(* IEC 61131-3 sources: Test-Git_ESME26/TestProgettoESME_26.fbsproj/PacDriveLib Migration/Motion/Homing (part 2) *)

(* ---- PDL_FB_HomeSetPos.fb.st ---- *)
FUNCTION_BLOCK PDL_FB_HomeSetPos
VAR_INPUT
	i_xEnable             : BOOL;
	i_ifDrive             : MOIN.IF_Axis;
	i_etMode              : PDL_ET_HomeSetPosMode;
	i_lrHomePosition      : LREAL;
	i_lrEncoderPosition   : LREAL;
	i_lrAbsEncOffset      : LREAL;
	i_lrUserPeriod        : LREAL;
	i_lrRestoreWindow     : LREAL;
	i_pstRestorePosRetain : POINTER TO PDL_ST_AxisRestorePosition;
	i_xExecute            : BOOL;
	iq_lencEncoder        : MOIN.IF_LogicalEncoder;
END_VAR
VAR_OUTPUT
	q_xActive           : BOOL;
	q_xReady            : BOOL;
	q_xBusy             : BOOL;
	q_xDone             : BOOL;
	q_etDiag            : GD.ET_Diag     := GD.ET_Diag.Ok;
	q_etDiagExt         : PDL_ET_DiagExt := PDL_ET_DiagExt.Disabled;
	q_sMsg              : STRING[80];
	q_lrPosition        : LREAL;
	q_lrEncoderPosition : LREAL;
	q_xHomeOk           : BOOL;
END_VAR
VAR
	xEnableFlag                                : BOOL;
	diState                                    : DINT;
	lrEncoderPeriode                           : LREAL;
	lrTurns                                    : LREAL;
	lrModuloPosition                           : LREAL;
	lrEncPosition                              : LREAL;
	xInterfacesInitialized                     : BOOL;
	xSuccess                                   : BOOL;
	etDiagTemp                                 : GD.ET_Diag := GD.ET_Diag.Ok;
	etDiagExtTemp                              : PDL_ET_DiagExt := PDL_ET_DiagExt.Ok;
	sDummyString                               : STRING[80];
	fbLoggerPoint                              : APL.FB_LoggerPoint;
	fbSetPosAxis                               : PLCO.MC_SetPosition;
	fbSetPosLenc                               : PLCO.MC_SetPosition;
	ifScalingAccess                            : DMFI.IF_ScalingAccess;
	ifScaling                                  : DMFI.IF_Scaling;
	ifGetParentDevice                          : DTSI.IF_GetParentDevice;
	ifDeviceAccess                             : DTSI.IF_DeviceAccess;
	ifEncoderAccess                            : DDI.IF_EncoderAccess;
	ifEncoder                                  : DDI.IF_Encoder;
	etModeOld                                  : PDL_ET_HomeSetPosMode;
	lrQuotientEncPeriodToUserPeriod            : LREAL;
	diTruncFromQuotient                        : DINT;
	lrAbsDifferenceQuotientToTruncFromQuotient : LREAL;
	xUserPeriodFitsIntoEncoderPeriod           : BOOL;
END_VAR

IF i_xEnable AND NOT xEnableFlag THEN (* Input action by rising edge of enable *)
	xEnableFlag := TRUE;
	THIS^.fbLoggerPoint.AddLogEntry(
		i_etLogLevel := APL.ET_LogLevel.UserAction, i_etDiag := q_etDiag, i_udiDiagExt := q_etDiagExt, i_sMessage := 'enable function block',
	);
	q_xActive              := TRUE;
	q_xReady               := FALSE;
	q_xBusy                := FALSE;
	q_xDone                := FALSE;
	q_xHomeOk              := FALSE;
	xInterfacesInitialized := Init_Interfaces();
	IF xInterfacesInitialized THEN
		etModeOld := i_etMode;
		q_xReady  := TRUE;
		SetDiagOutput(i_etDiag := GD.ET_Diag.OK, i_etDiagExt := PDL_ET_DiagExt.WaitForExecute, i_sMsg := '');
		diState := 10;
	END_IF
	i_ifDrive.xIsHomed := FALSE;

ELSIF NOT i_xEnable AND xEnableFlag THEN (* Output action by falling edge of enable *)
	xEnableFlag := FALSE;
	THIS^.fbLoggerPoint.AddLogEntry(
		i_etLogLevel := APL.ET_LogLevel.UserAction, i_etDiag := q_etDiag, i_udiDiagExt := q_etDiagExt, i_sMessage := 'disable function block',
	);
	xInterfacesInitialized := FALSE;
	q_xActive              := FALSE;
	q_xReady               := FALSE;
	q_xBusy                := FALSE;
	q_xDone                := FALSE;
	q_lrPosition           := 0.0;
	q_lrEncoderPosition    := 0.0;
	q_xHomeOk              := FALSE;
	SetDiagOutput(i_etDiag := GD.ET_Diag.Ok, i_etDiagExt := PDL_ET_DiagExt.Disabled, i_sMsg := '');
	diState := 0;
ELSIF NOT q_xActive THEN
	RETURN;
END_IF

IF xInterfacesInitialized THEN
	q_lrPosition        := i_ifDrive.RefPosition;
	IF iq_lencEncoder <> 0 THEN
		q_lrEncoderPosition := iq_lencEncoder.RefPosition;
	ELSE
		q_lrEncoderPosition := 0;
	END_IF
	q_xBusy             := q_etDiag = GD.ET_Diag.Ok AND NOT q_xDone AND diState > 10;
ELSE
	diState  := 0;
	q_xReady := FALSE;
	RETURN;
END_IF

CASE diState OF
	0: (* Idle *)
		;
	10: (* wait for xExecute *)
		IF i_xExecute THEN
			IF etModeOld <> i_etMode THEN
				etModeOld              := i_etMode;
				xInterfacesInitialized := Init_Interfaces();
			END_IF
			lrEncoderPeriode := 0;

			THIS^.fbLoggerPoint.AddLogEntry(
				i_etLogLevel := APL.ET_LogLevel.UserAction,
				i_etDiag     := q_etDiag,
				i_udiDiagExt := q_etDiagExt,
				i_sMessage   := 'start homing',
				q_etDiag     =>,
				q_etDiagExt  =>
			);

			lrEncoderPeriode 			:= ifEncoder.Revolutions
											* ifScaling.PositionResolution
											* TO_LREAL(ifScaling.GearIn) / TO_LREAL(ifScaling.GearOut)
											* TO_LREAL( ifEncoder.GearOut) / TO_LREAL(ifEncoder.GearIn);

						// Calculation if UserPeriod fits into EncoderPeriod
			IF (i_lrUserPeriod > CMT.Gc_lrZeroTolerance) AND (lrEncoderPeriode > CMT.Gc_lrZeroTolerance) THEN

				lrQuotientEncPeriodToUserPeriod					:= lrEncoderPeriode/i_lrUserPeriod;
				diTruncFromQuotient 							:= TRUNC(lrQuotientEncPeriodToUserPeriod);
				lrAbsDifferenceQuotientToTruncFromQuotient		:= ABS (lrQuotientEncPeriodToUserPeriod - TO_LREAL(diTruncFromQuotient));

				IF (lrAbsDifferenceQuotientToTruncFromQuotient < CMT.Gc_lrZeroTolerance)
				OR ((1 - lrAbsDifferenceQuotientToTruncFromQuotient < CMT.Gc_lrZeroTolerance) AND (lrAbsDifferenceQuotientToTruncFromQuotient <= 1)) THEN
					xUserPeriodFitsIntoEncoderPeriod	:= TRUE;
				ELSE
					xUserPeriodFitsIntoEncoderPeriod	:= FALSE;
				END_IF

			END_IF

			CASE i_etMode OF
				//---------------------------------------
				PDL_ET_HomeSetPosMode.RestorePosFromRetain,
				PDL_ET_HomeSetPosMode.SetPosAxisPosition,
				PDL_ET_HomeSetPosMode.SetPosLogEncoderPosition,
				PDL_ET_HomeSetPosMode.SetPosAxisAndLogEncoderPosition,
				PDL_ET_HomeSetPosMode.RestorePosFromAxisencoder:
					//---------------------------------------

					//Input-Parameter-Checks
					IF i_etMode = PDL_ET_HomeSetPosMode.RestorePosFromAxisEncoder OR i_etMode = PDL_ET_HomeSetPosMode.RestorePosFromRetain THEN
						IF (ABS(ifEncoder.Revolutions) < 1.0E-3) THEN
							SetDiagOutput(	i_etDiag := GD.ET_Diag.DriveConditionInvalid,
											i_etDiagExt := PDL_ET_DiagExt.DriveEncoderInvalid,
											i_sMsg := ''
							);
							diState := 0;
							RETURN;
						END_IF

						IF (i_lrUserPeriod < 0.0) THEN
							SetDiagOutput(
								i_etDiag    := GD.ET_Diag.InputParameterInvalid,
								i_etDiagExt := PDL_ET_DiagExt.UserPeriodRange,
								i_sMsg      := '0.0 <= i_lrUserPeriod'
							);
							diState := 0;
							RETURN;
							// if UserPeriod = 0: Check if AbsEncOffset > 0
						ELSIF
							i_etMode = PDL_ET_HomeSetPosMode.RestorePosFromAxisencoder AND
							(i_lrUserPeriod = 0.0) AND
							((i_lrAbsEncOffset < 0) OR (i_lrAbsEncOffset > lrEncoderPeriode))
						THEN
							SetDiagOutput(
								i_etDiag    := GD.ET_Diag.InputParameterInvalid,
								i_etDiagExt := PDL_ET_DiagExt.AbsEncOffsetRange,
								i_sMsg      := STANDARD.CONCAT('0.0 < i_lrAbsEncOffset <= ', SE_CTBX.FC_LrealToString(i_sFormat := '#0.00', i_lrInput := lrEncoderPeriode))
							);
							diState := 0;
							RETURN;
							// Check if UserPeriode fits into EncoderPeriode
						ELSIF i_etMode = PDL_ET_HomeSetPosMode.RestorePosFromAxisencoder AND (i_lrUserPeriod > 0.0) AND NOT xUserPeriodFitsIntoEncoderPeriod
						THEN
							SetDiagOutput(
								i_etDiag    := GD.ET_Diag.InputParameterInvalid,
								i_etDiagExt := PDL_ET_DiagExt.UserPeriodRange,
								i_sMsg      := STANDARD.CONCAT('i_lrUserPeriod has to be a divsior of ',SE_CTBX.FC_LrealToString(i_sFormat := '#0.00', i_lrInput := lrEncoderPeriode))
							);
							diState := 0;
							RETURN;
						END_IF
					END_IF

					q_xHomeOk := FALSE;
					q_xBusy   := TRUE;
					q_xDone   := FALSE;
					SetDiagOutput(i_etDiag := GD.ET_Diag.Ok, i_etDiagExt := PDL_ET_DiagExt.WaitUntilHomingDone, i_sMsg := '');
					diState := 20;
				ELSE
					SetDiagOutput(i_etDiag := GD.ET_Diag.InputParameterInvalid, i_etDiagExt := PDL_ET_DiagExt.UnknownMode, i_sMsg := '');
					diState := 0;
			END_CASE
		END_IF
	20:
		CASE i_etMode OF
			//---------------------------------------
			PDL_ET_HomeSetPosMode.RestorePosFromRetain: (* Restore axis position from stored and actual Values of position and encoder position *)
				//---------------------------------------
				IF i_pstRestorePosRetain > 0 THEN
					PDL_FC_RestoreAxisPosition(
						i_ifDrive           := i_ifDrive,
						i_lrUserPeriod      := i_lrUserPeriod,
						i_lrRestoreWindow   := i_lrRestoreWindow,
						i_stRestorePosition := i_pstRestorePosRetain^,
						q_etDiag            => etDiagTemp,
						q_etDiagExt         => etDiagExtTemp,
						q_sMsg              => sDummyString
					);
					IF etDiagTemp = GD.ET_Diag.Ok THEN
						diState := 30;
					ELSE
						CASE etDiagExtTemp OF
							PDL_ET_DiagExt.CheckSumInvalid:
								SetDiagOutput(
									i_etDiag    := GD.ET_Diag.InputParameterInvalid,
									i_etDiagExt := PDL_ET_DiagExt.CheckSumInvalid,
									i_sMsg      := 'FB_HomeSetPos: FC_RestoreAxisPosition'
								);
							PDL_ET_DiagExt.DataNVRamInvalid:
								SetDiagOutput(
									i_etDiag    := GD.ET_Diag.InputParameterInvalid,
									i_etDiagExt := PDL_ET_DiagExt.DataNVRamInvalid,
									i_sMsg      := 'FB_HomeSetPos: FC_RestoreAxisPosition'
								);
							PDL_ET_DiagExt.SercosNotInPhaseFour:
								SetDiagOutput(
									i_etDiag    := GD.ET_Diag.DriveConditionInvalid,
									i_etDiagExt := PDL_ET_DiagExt.SercosNotInPhaseFour,
									i_sMsg      := 'FB_HomeSetPos: FC_RestoreAxisPosition'
								);
							PDL_ET_DiagExt.DriveEncoderInvalid:
								SetDiagOutput(
									i_etDiag    := GD.ET_Diag.DriveConditionInvalid,
									i_etDiagExt := PDL_ET_DiagExt.DriveEncoderInvalid,
									i_sMsg      := 'FB_HomeSetPos: FC_RestoreAxisPosition'
								);
							PDL_ET_DiagExt.OutOfRestoreWindow:
								SetDiagOutput(
									i_etDiag    := GD.ET_Diag.LimitReached,
									i_etDiagExt := PDL_ET_DiagExt.OutOfRestoreWindow,
									i_sMsg      := 'FB_HomeSetPos: FC_RestoreAxisPosition'
								);
							PDL_ET_DiagExt.UnexpectedFeedback:
								SetDiagOutput(
									i_etDiag    := GD.ET_Diag.UnexpectedProgramBehavior,
									i_etDiagExt := PDL_ET_DiagExt.UnexpectedFeedback,
									i_sMsg      := Standard.CONCAT('FB_HomeSetPos: FC_RestoreAxisPosition: ', sDummyString)
								);
							PDL_ET_DiagExt.RestoreInterrupted:
								SetDiagOutput(
									i_etDiag    := GD.ET_Diag.DriveConditionInvalid,
									i_etDiagExt := PDL_ET_DiagExt.RestoreInterrupted,
									i_sMsg      := 'FB_HomeSetPos: FC_RestoreAxisPosition'
								);
						END_CASE
						diState := 0;
					END_IF
				ELSE
					SetDiagOutput(
						i_etDiag := GD.ET_Diag.InputParameterInvalid, i_etDiagExt := PDL_ET_DiagExt.PointerRestorePosRetainInvalid, i_sMsg := ''
					);
					diState := 0;
				END_IF
				//-------------------------------------
			PDL_ET_HomeSetPosMode.SetPosAxisPosition:
				//-------------------------------------

				THIS^.fbSetPosAxis(Axis := i_ifDrive, Execute := TRUE, Position := i_lrHomePosition, Relative := FALSE);

				IF THIS^.fbSetPosAxis.Done THEN
					diState := 30;
				ELSIF THIS^.fbSetPosAxis.Error THEN
					SetDiagOutput(
						i_etDiag    := GD.ET_Diag.UnexpectedProgramBehavior,
						i_etDiagExt := PDL_ET_DiagExt.UnexpectedFeedback,
						i_sMsg      := CONCAT('MC_Setposition.ErrorID: ', PLCO.FC_EtResultToString(THIS^.fbSetPosAxis.ErrorId))
					);
					THIS^.fbSetPosAxis(Execute := FALSE);
					diState := 0;
				END_IF

				//-------------------------------------------
			PDL_ET_HomeSetPosMode.SetPosLogEncoderPosition:
				//-------------------------------------------
				THIS^.fbSetPosLenc(Axis := iq_lencEncoder, Execute := TRUE, Position := i_lrEncoderPosition, Relative := FALSE);

				IF THIS^.fbSetPosLenc.Done THEN
					diState := 30;
				ELSIF THIS^.fbSetPosLenc.Error THEN
					SetDiagOutput(
						i_etDiag    := GD.ET_Diag.UnexpectedProgramBehavior,
						i_etDiagExt := PDL_ET_DiagExt.UnexpectedFeedback,
						i_sMsg      := CONCAT('MC_Setposition.ErrorID: ', PLCO.FC_EtResultToString(THIS^.fbSetPosLenc.ErrorId))
					);
					THIS^.fbSetPosLenc(Execute := FALSE);
					diState := 0;
				END_IF

				//--------------------------------------------------
			PDL_ET_HomeSetPosMode.SetPosAxisAndLogEncoderPosition:
				//--------------------------------------------------
				THIS^.fbSetPosLenc(Axis := iq_lencEncoder, Execute := TRUE, Position := i_lrEncoderPosition, Relative := FALSE);

				THIS^.fbSetPosAxis(Axis := i_ifDrive, Execute := TRUE, Position := i_lrHomePosition, Relative := FALSE);

				IF THIS^.fbSetPosAxis.Done AND THIS^.fbSetPosLenc.Done THEN
					diState := 30;
				ELSIF THIS^.fbSetPosAxis.Error THEN
					SetDiagOutput(
						i_etDiag    := GD.ET_Diag.UnexpectedProgramBehavior,
						i_etDiagExt := PDL_ET_DiagExt.UnexpectedFeedback,
						i_sMsg      := CONCAT('MC_Setposition.ErrorID: ', PLCO.FC_EtResultToString(THIS^.fbSetPosAxis.ErrorId))
					);
					THIS^.fbSetPosAxis(Execute := FALSE);
					THIS^.fbSetPosLenc(Execute := FALSE);
					diState := 0;

				ELSIF THIS^.fbSetPosLenc.Error THEN
					SetDiagOutput(
						i_etDiag    := GD.ET_Diag.UnexpectedProgramBehavior,
						i_etDiagExt := PDL_ET_DiagExt.UnexpectedFeedback,
						i_sMsg      := CONCAT('MC_Setposition.ErrorID: ', PLCO.FC_EtResultToString(THIS^.fbSetPosLenc.ErrorId))
					);
					THIS^.fbSetPosLenc(Execute := FALSE);
					THIS^.fbSetPosAxis(Execute := FALSE);
					diState := 0;
				END_IF

				//--------------------------------------------
			PDL_ET_HomeSetPosMode.RestorePosFromAxisencoder: (* Gebertyp feststellen und GeberPeriode berechnen *)
				//--------------------------------------------
				lrTurns          := ifEncoder.Revolutions;
				IF NOT ifScaling.InvertDirection THEN (* motor direction right *)
					lrEncPosition := ifEncoder.Position;
				ELSE
					lrEncPosition := lrEncoderPeriode - ifEncoder.Position;
				END_IF
				(* In a round axis, position is always within the user period, AbsEncOffset is not allowed *)
				IF i_lrUserPeriod > 0.0 THEN
					lrModuloPosition := lrEncPosition - TRUNC_INT(lrEncPosition / i_lrUserPeriod) * i_lrUserPeriod;
					THIS^.fbSetPosAxis(Axis := i_ifDrive, Execute := TRUE, Position := lrModuloPosition, Relative := FALSE);
				ELSE
					(* Absolute axis *)
					(*---------------*)
					(* The range of the encoder period is between 0 and encoder period *)
					(* In absolute systems it makes sense to have an Offset to have neg. positions *)
					(* Of course, the Offset reduces the upper limit of the max. travel *)

					(* without AbsEncOffset *)
					(* 		   +---------------------------------------------------------------------------------------------------+ 	                   	*)
					(*         0                                                                                                EncoderPeriode				*)

					(* with AbsEncOffset *)
					(* 		   +---------------------+-----------------------------------------------------------------------------+ 	                   	*)
					(*		-AbsEncOffset			0												                   EncoderPeriode - AbsEncOffset		*)
					IF (lrEncPosition > (lrEncoderPeriode - i_lrAbsEncOffset)) THEN
						THIS^.fbSetPosAxis(Axis := i_ifDrive, Execute := TRUE, Position := lrEncPosition - lrEncoderPeriode, Relative := FALSE);
					ELSE
						THIS^.fbSetPosAxis(Axis := i_ifDrive, Execute := TRUE, Position := lrEncPosition, Relative := FALSE);
					END_IF
				END_IF
				IF THIS^.fbSetPosAxis.Done THEN
					diState := 30;
				ELSE
					SetDiagOutput(
						i_etDiag    := GD.ET_Diag.UnexpectedProgramBehavior,
						i_etDiagExt := PDL_ET_DiagExt.UnexpectedFeedback,
						i_sMsg      := CONCAT('MC_Setposition.ErrorID: ', PLCO.FC_EtResultToString(THIS^.fbSetPosAxis.ErrorId))
					);
					THIS^.fbSetPosAxis(Execute := FALSE);
					diState := 0;
				END_IF
			ELSE (* End case mode / Home.Mode unknown *)
				SetDiagOutput(i_etDiag := GD.ET_Diag.InputParameterInvalid, i_etDiagExt := PDL_ET_DiagExt.UnknownMode, i_sMsg := '');
				diState := 0;
		END_CASE
	30: (* Set Outputs for Homing Results *)
		SetDiagOutput(i_etDiag := GD.ET_Diag.Ok, i_etDiagExt := PDL_ET_DiagExt.HomingDone, i_sMsg := '');
		q_xHomeOK := TRUE;
		q_xDone   := TRUE;
		THIS^.fbSetPosAxis(Execute := FALSE);
		THIS^.fbSetPosLenc(Execute := FALSE);
		diState := 40;
	40: (* Wait for NOT Execute *)
		IF NOT i_xExecute THEN
			SetDiagOutput(i_etDiag := GD.ET_Diag.Ok, i_etDiagExt := PDL_ET_DiagExt.WaitForExecute, i_sMsg := '');
			diState := 10;
		END_IF
	ELSE (* End of case *)
		SetDiagOutput(
			i_etDiag := GD.ET_Diag.UnexpectedProgramBehavior, i_etDiagExt := PDL_ET_DiagExt.UnknownState, i_sMsg := DINT_TO_STRING(diState)
		);
		diState := 0;
END_CASE

(* ---- PDL_FB_HomeTorque.fb.st ---- *)
FUNCTION_BLOCK PDL_FB_HomeTorque
VAR_INPUT
	i_xEnable        : BOOL;
	i_ifDrive        : MOIN.IF_Axis;
	i_lrMaxTorque    : LREAL;
	i_diTorqueTime   : DINT;
	i_lrLowLimit     : LREAL;
	i_lrHighLimit    : LREAL;
	i_etMode         : PDL_ET_HomeTorqueMode;
	i_lrOffset       : LREAL;
	i_lrMaxTravel    : LREAL;
	i_lrHomePosition : LREAL;
	i_lrVel          : LREAL;
	i_lrAcc          : LREAL;
	i_lrDec          : LREAL;
	i_lrJerk         : LREAL;
	i_xStart         : BOOL;
END_VAR
VAR_OUTPUT
	q_xActive                  : BOOL;
	q_xReady                   : BOOL;
	q_etDiag                   : GD.ET_Diag := GD.ET_Diag.Ok;
	q_etDiagExt                : PDL_ET_DiagExt := PDL_ET_DiagExt.Disabled;
	q_sMsg                     : STRING[80];
	q_xMotionInstructionActive : BOOL;
	q_lrPosition               : LREAL;
	q_xHomeOk                  : BOOL;
END_VAR
VAR
	fbLoggerPoint            : APL.FB_LoggerPoint;
	ifDeviceTreeObjectAccess : UFMPLCI.IF_DeviceTreeObjectAccess;
	sDriveName               : STRING(80);
	ifDriveConfigAccess      : DDI.IF_DriveConfigAccess;
	ifDriveConfig            : DDI.IF_DriveConfig;
	ifDriveCurrent           : DDI.IF_DriveCurrent;
	ifDriveCurrentAccess     : DDI.IF_DriveCurrentAccess;
	ifDrive2                 : DDI.IF_Drive2;
	ifDrive2Access           : DDI.IF_Drive2Access;
	ifDriveAccess            : DMFI.IF_DriveAccess;
	ifDrive                  : DMFI.IF_Drive;
	xSuccess                 : BOOL;
	xInterfacesInitialised   : BOOL;

	xEnableFlag : BOOL;

	diState   : DINT;
	etDiagExt : PDL_ET_DiagExt;

	fbStop                      : PLCO.MC_Stop;
	fbSetPos                    : PLCO.MC_SetPosition;
	xError                      : BOOL;
	etResult                    : SE_Async.ET_Result;
	sResultMsg                  : STRING(80);
	xStartFlag                  : BOOL;
	lrOldUserCurrentLimit       : REAL;
	lrOldTrackingDeviationLimit : LREAL;
	fbSetTrackDev               : PDL_FB_SetTrackingDeviation;
	fbResetTrackDev             : PDL_FB_ResetTrackingDeviation;
	fbPosOnTorque               : PDL_FB_PosOnTorque;
END_VAR

IF i_xEnable AND NOT xEnableFlag THEN
	xEnableFlag := TRUE;
	THIS^.fbLoggerPoint.AddLogEntry(
		i_etLogLevel := APL.ET_LogLevel.UserAction,
		i_etDiag     := q_etDiag,
		i_udiDiagExt := q_etDiagExt,
		i_sMessage   := 'enable function block',
		q_etDiag     =>,
		q_etDiagExt  =>
	);
	q_xActive                  := TRUE;
	q_xReady                   := FALSE;
	q_xHomeOk                  := FALSE;
	q_xMotionInstructionActive := FALSE;
	diState                    := 0;
	SetDiagOutput(
		i_etDiag    := GD.ET_Diag.OK,
		i_etDiagExt := PDL_ET_DiagExt.Initializing,
		i_sMsg      := ''
	);

	xSuccess := InitInterfaces();
	IF NOT xSuccess THEN
		xInterfacesInitialised := FALSE;
		RETURN;
	END_IF

	xSuccess := InputParameterCheck();
	IF NOT xSuccess THEN
		RETURN;
	END_IF
	i_ifDrive.xIsHomed         := FALSE;
	fbStop(Execute := FALSE);

	xStartFlag             := FALSE;
	xInterfacesInitialised := TRUE;
	lrOldUserCurrentLimit  := ifDriveCurrent.UserCurrentLimit;
	diState                := -10000;

ELSIF NOT i_xEnable AND xEnableFlag THEN
	xEnableFlag := FALSE;
	THIS^.fbLoggerPoint.AddLogEntry(
		i_etLogLevel := APL.ET_LogLevel.UserAction,
		i_etDiag     := q_etDiag,
		i_udiDiagExt := q_etDiagExt,
		i_sMessage   := 'disable function block',
		q_etDiag     =>,
		q_etDiagExt  =>
	);
	q_xReady := FALSE;
	IF xInterfacesInitialised THEN
		IF ABS(ifDrive2.TrackingDeviation) > lrOldTrackingDeviationLimit THEN
			fbSetPos(
				Execute  := TRUE,
				Position := ifDrive.ActualPosition,
				Relative := FALSE
			);
			fbSetPos(Execute := FALSE);
		END_IF
		SetDiagOutput(
			i_etDiag    := GD.ET_Diag.OK,
			i_etDiagExt := PDL_ET_DiagExt.WaitUntilDisabled,
			i_sMsg      := ''
		);
		ifDriveCurrent.UserCurrentLimit := lrOldUserCurrentLimit;
		diState                         := -10010;
	ELSE
		q_xActive                  := FALSE;
		q_lrPosition               := 0.0;
		q_xMotionInstructionActive := FALSE;
		q_xHomeOk                  := FALSE;
		xInterfacesInitialised     := FALSE;
		SetDiagOutput(
			i_etDiag    := GD.ET_Diag.OK,
			i_etDiagExt := PDL_ET_DiagExt.Disabled,
			i_sMsg      := ''
		);
		diState := 0;
	END_IF
END_IF

IF xInterfacesInitialised AND q_xActive THEN
	IF i_ifDrive.etAxisState < MOIN.ET_AxisState.Standstill AND diState > 0 AND diState < 100 THEN
		diState                    := 0;
		q_xReady                   := FALSE;
		q_xMotionInstructionActive := FALSE;
		SetDiagOutput(
			i_etDiag    := GD.ET_Diag.DriveConditionInvalid,
			i_etDiagExt := PDL_ET_DiagExt.DriveNotReady,
			i_sMsg 		:= STANDARD.CONCAT(sDriveName,': AxisState < Standstill')
		);
	END_IF
	q_lrPosition := i_ifDrive.RefPosition;
END_IF

CASE diState OF
	-10000: // State for Set TrackingDeviation
		IF SE_Async.G_ifAsyncMgr.xInitDone THEN
			fbSetTrackDev.ifDrive2 := ifDrive2;
			SE_Async.G_ifAsyncMgr.Start(
				i_ifAsync    := fbSetTrackDev,
				q_etResult   => etResult,
				q_sResultMsg => sResultMsg,
				q_xError     => xError
			);
			IF xError THEN
				AsyncExtDiagTranslation(i_etResult := etResult);
				RETURN;
			ELSE
				diState := -10001;
			END_IF
		ELSE
			SE_Async.G_ifAsyncMgr.Init(
				q_xError     => xError,
				q_etResult   => etResult,
				q_sResultMsg => sResultMsg
			);
			IF xError THEN
				AsyncExtDiagTranslation(i_etResult := etResult);
				diState := 0;
			END_IF
		END_IF
	-10001: //Waiting State for Set TrackingDeviation Done
		IF fbSetTrackDev.xDone THEN
			lrOldTrackingDeviationLimit := fbSetTrackDev.lrOldTrackDevLim;
			q_xReady                    := TRUE;
			SetDiagOutput(
				i_etDiag    := GD.ET_Diag.OK,
				i_etDiagExt := PDL_ET_DiagExt.WaitForStart,
				i_sMsg      := ''
			);
			diState := 10;
		END_IF
	-10010:
		IF SE_Async.G_ifAsyncMgr.xInitDone THEN
			fbResetTrackDev.ifDrive2         := ifDrive2;
			fbResetTrackDev.lrOldTrackDevLim := lrOldTrackingDeviationLimit;
			SE_Async.G_ifAsyncMgr.Start(
				i_ifAsync    := fbResetTrackDev,
				q_etResult   => etResult,
				q_sResultMsg => sResultMsg,
				q_xError     => xError
			);
			IF xError THEN
				AsyncExtDiagTranslation(i_etResult := etResult);
				RETURN;
			ELSE
				diState := -10011;
			END_IF
		ELSE
			SE_Async.G_ifAsyncMgr.Init(
				q_xError     => xError,
				q_etResult   => etResult,
				q_sResultMsg => sResultMsg
			);
			IF xError THEN
				AsyncExtDiagTranslation(i_etResult := etResult);
				diState := 0;
			END_IF
		END_IF
	-10011: // Wait for TrackDev reset
		IF fbResetTrackDev.xDone THEN
			fbStop(Execute := TRUE);
			diState := 100;
		END_IF
	0: (* Exception or No Enable or ready  *)
		;
	10: (* Wait for Start*)
		IF i_xStart AND NOT xStartFlag THEN
			xStartFlag := TRUE;
			THIS^.fbLoggerPoint.AddLogEntry(
				i_etLogLevel := APL.ET_LogLevel.UserAction,
				i_etDiag     := q_etDiag,
				i_udiDiagExt := q_etDiagExt,
				i_sMessage   := 'start homing'
			);
			xSuccess := InputParameterCheck();
			IF NOT xSuccess THEN
				q_xReady := FALSE;
				diState  := 0;
				RETURN;
			END_IF
			q_xHomeOk          := FALSE;
			i_ifDrive.xIsHomed := FALSE;

			CASE i_etMode OF
				PDL_ET_HomeTorqueMode.PosDirectionMaxTorque: (* Mode 0:  pos. Direction and MaxTorque *)
					fbPosOnTorque(
						i_ifDrive        := i_ifDrive,
						i_lrMaxTorque    := i_lrMaxTorque,
						i_diTorqueTime   := i_diTorqueTime,
						i_lrLowLimit     := i_lrLowLimit,
						i_lrHighLimit    := i_lrHighLimit,
						i_lrMaxTravel    := ABS(i_lrMaxTravel),
						i_lrOffset       := -ABS(i_lrOffset),
						i_lrVelocity     := i_lrVel,
						i_lrAcceleration := i_lrAcc,
						i_lrDeceleration := i_lrDec,
						i_lrJerk         := i_lrJerk,
						i_xStart         := TRUE
					);
				PDL_ET_HomeTorqueMode.NegDirectionMaxTorque: (* Mode 1:  neg. Direction and MaxTorque *)
					fbPosOnTorque(
						i_ifDrive        := i_ifDrive,
						i_lrMaxTorque    := i_lrMaxTorque,
						i_diTorqueTime   := i_diTorqueTime,
						i_lrLowLimit     := i_lrLowLimit,
						i_lrHighLimit    := i_lrHighLimit,
						i_lrMaxTravel    := -ABS(i_lrMaxTravel),
						i_lrOffset       := ABS(i_lrOffset),
						i_lrVelocity     := i_lrVel,
						i_lrAcceleration := i_lrAcc,
						i_lrDeceleration := i_lrDec,
						i_lrJerk         := i_lrJerk,
						i_xStart         := TRUE
					);
				ELSE
					q_xReady := FALSE;
					SetDiagOutput(
						i_etDiag    := GD.ET_Diag.InputParameterInvalid,
						i_etDiagExt := PDL_ET_DiagExt.UnknownMode,
						i_sMsg      := ''
					);
					diState := 0;
					RETURN;
			END_CASE
			q_xMotionInstructionActive := TRUE;
			SetDiagOutput(
				i_etDiag    := GD.ET_Diag.OK,
				i_etDiagExt := PDL_ET_DiagExt.WaitUntilMaxTorqueReached,
				i_sMsg      := ''
			);
			diState := 20;
		ELSIF NOT i_xStart AND xStartFlag THEN
			xStartFlag := FALSE;
		END_IF
	20:
		fbPosOnTorque(i_xStart := FALSE);
		IF fbPosOnTorque.q_etDiagExt = PDL_ET_DiagExt.WaitForStart THEN
			q_xHomeOk                  := fbPosOnTorque.q_xTorqueOk;
			q_xMotionInstructionActive := FALSE;
			IF q_xHomeOk THEN
				fbSetpos(
					Execute  := TRUE,
					Relative := FALSE,
					Position := i_lrHomePosition
				);
				IF fbSetpos.Error THEN
					SetDiagOutput(
						i_etDiag    := GD.ET_Diag.UnexpectedProgramBehavior,
						i_etDiagExt := PDL_ET_DiagExt.UnexpectedFeedback,
						i_sMsg      := CONCAT('MC_Setpos: ',PLCO.FC_EtResultToString(fbSetpos.ErrorId))
					);
					RETURN;
				END_IF
				SetDiagOutput(
					i_etDiag    := GD.ET_Diag.OK,
					i_etDiagExt := PDL_ET_DiagExt.HomingDone,
					i_sMsg      := ''
				);
				fbSetpos(Execute := FALSE);
				diState := 10;
			ELSE
				i_ifDrive.xIsHomed := FALSE;
				q_xReady           := FALSE;
				SetDiagOutput(
					i_etDiag    := GD.ET_Diag.UnexpectedProgramBehavior,
					i_etDiagExt := PDL_ET_DiagExt.UnexpectedFeedback,
					i_sMsg      := CONCAT('FB_PosOnTorque: ',PDL_FC_EtDiagExtToString(i_etDiagExt := fbPosOnTorque.q_etDiagExt))
				);
				diState := 0;
			END_IF

		ELSIF fbPosOnTorque.q_etDiag <> GD.ET_Diag.Ok THEN
			i_ifDrive.xIsHomed         := FALSE;
			q_xMotionInstructionActive := FALSE;
			q_xReady                   := FALSE;
			SetDiagOutput(
				i_etDiag    := fbPosOnTorque.q_etDiag,
				i_etDiagExt := fbPosOnTorque.q_etDiagExt,
				i_sMsg      := fbPosOnTorque.q_sMsg
			);
			diState := 0;
		END_IF
	100: (* Wait until stopped *)
		fbStop(Execute := TRUE);
		IF
			i_ifDrive.etAxisState = MOIN.ET_AxisState.Disabled OR
			i_ifDrive.etAxisState = MOIN.ET_AxisState.ErrorStop OR
			i_ifDrive.etAxisState = MOIN.ET_AxisState.Standstill OR
			fbStop.Done
		THEN
			fbStop(Execute := FALSE);
			xInterfacesInitialised     := FALSE;
			q_xMotionInstructionActive := FALSE;
			q_xActive                  := FALSE;
			q_lrPosition               := 0.0;
			q_xHomeOk                  := FALSE;

			SetDiagOutput(
				i_etDiag    := GD.ET_Diag.OK,
				i_etDiagExt := PDL_ET_DiagExt.Disabled,
				i_sMsg      := ''
			);
			diState := 0;
		END_IF

		IF fbStop.Error AND fbStop.ErrorId <> PLCO.ET_Result.StoppingInterrupted THEN
			q_xMotionInstructionActive := FALSE;
			q_xReady                   := FALSE;
			SetDiagOutput(
				i_etDiag    := GD.ET_Diag.UnexpectedProgramBehavior,
				i_etDiagExt := PDL_ET_DiagExt.UnexpectedFeedback,
				i_sMsg      := CONCAT('MC_Stop: ',PLCO.FC_EtResultToString(fbStop.ErrorId))
			);
			fbStop(Execute := FALSE);
			diState := 0;
		END_IF

		(* Ende Case *)
	ELSE
		q_xReady                   := FALSE;
		q_xMotionInstructionActive := FALSE;
		SetDiagOutput(
			i_etDiag    := GD.ET_Diag.UnexpectedProgramBehavior,
			i_etDiagExt := PDL_ET_DiagExt.UnknownState,
			i_sMsg      := DINT_TO_STRING(diState)
		);
		diState := 0;
END_CASE

(* ---- PDL_FB_HomeTp.fb.st ---- *)
FUNCTION_BLOCK PDL_FB_HomeTp
VAR_INPUT
	i_xEnable         : BOOL;
	i_ifDrive         : MOIN.IF_Axis;
	i_ifTouchProbe    : PLCO.MC_Trigger_Ref;
	i_etMode          : PDL_ET_HomeTpMode;
	i_lrOffset        : LREAL;
	i_lrMaxTravel     : LREAL;
	i_lrHomePosition  : LREAL;
	i_lrVel           : LREAL;
	i_lrAcc           : LREAL;
	i_lrDec           : LREAL;
	i_lrJerk          : LREAL;
	i_xHwLimitNeg     : BOOL;
	i_xHwLimitPos     : BOOL;
	i_xRotativeSystem : BOOL;
	i_xStart          : BOOL;
END_VAR
VAR_OUTPUT
	q_xActive                  : BOOL;
	q_xReady                   : BOOL;
	q_etDiag                   : GD.ET_Diag := GD.ET_Diag.Ok;
	q_etDiagExt                : PDL_ET_DiagExt := PDL_ET_DiagExt.Disabled;
	q_sMsg                     : STRING[80];
	q_xMotionInstructionActive : BOOL;
	q_lrPosition               : LREAL;
	q_xHomeOk                  : BOOL;
END_VAR
VAR
	xEnableFlag   : BOOL;
	diState       : DINT;
	fbLoggerPoint : APL.FB_LoggerPoint;

	xLimitGivenDirection       : BOOL;
	xLimitGivenDirectionOld    : BOOL;
	xLimitOpposideDirection    : BOOL;
	xLimitOpposideDirectionOld : BOOL;
	lrDistance                 : LREAL;
	xMotionJobStarted          : BOOL;
	ifDeviceTreeObjectAccess   : UFMPLCI.IF_DeviceTreeObjectAccess;
	sDriveName                 : STRING(80);
	ifScalingAccess            : DMFI.IF_ScalingAccess;
	ifScaling                  : DMFI.IF_Scaling;
	ifDrive2Access             : DDI.IF_Drive2Access;
	ifDrive2                   : DDI.IF_Drive2;
	ifDriveAccess              : DMFI.IF_DriveAccess;
	ifDrive                    : DMFI.IF_Drive;
	ifDriveConfigAccess        : DDI.IF_DriveConfigAccess;
	ifDriveConfig              : DDI.IF_DriveConfig;
	ifTouprobeData             : IODI.IF_TouchprobeData;
	ifTouprobeDataAccess       : IODI.IF_TouchprobeDataAccess;
	fbTouchProbe               : PLCO.MC_TouchProbe;
	fbAbortTouchprobe          : PLCO.MC_AbortTrigger;
	fbStop                     : PLCO.MC_Stop;
	fbHalt                     : PLCO.MC_Halt;
	fbMoveAbsolute             : PLCO.MC_MoveAbsolute;
	fbMoveRelative             : PLCO.MC_MoveRelative;
	fbSetPos                   : PLCO.MC_SetPosition;

END_VAR

IF i_xEnable AND NOT xEnableFlag AND (diState = 0) THEN
	// detect positive flank on i_xEnable if FB is disabled
	xEnableFlag := TRUE;
	fbLoggerPoint.AddLogEntry(
		i_etLogLevel := APL.ET_LogLevel.UserAction, i_etDiag := q_etDiag, i_udiDiagExt := q_etDiagExt, i_sMessage := 'enable function block'
	);
	q_xActive                  := TRUE;
	q_xReady                   := FALSE;
	q_xMotionInstructionActive := FALSE;
	q_xHomeOk                  := FALSE;
	IF THIS^.EnableParameterCheck() THEN
		i_ifDrive.xIsHomed         := FALSE;
		fbStop(Execute := FALSE);
		fbSetPos(Execute := FALSE);
		fbAbortTouchprobe(Execute := FALSE);
		fbTouchProbe(Execute := FALSE);
		fbMoveAbsolute(Execute := FALSE);
		fbMoveRelative(Execute := FALSE);
		fbAbortTouchprobe.Axis := i_ifDrive;
		fbAbortTouchprobe.ifTrigger := i_ifTouchProbe;
		fbAbortTouchprobe(Execute := TRUE);
		IF fbAbortTouchprobe.Error THEN
			SetDiagOutput(
				i_etDiag    := GD.ET_Diag.UnexpectedProgramBehavior,
				i_etDiagExt := PDL_ET_DiagExt.UnexpectedFeedback,
				i_sMsg      := CONCAT('MC_AbortTrigger: ', PLCO.FC_EtResultToString(fbAbortTouchprobe.ErrorId))
			);
		ELSE
			q_xReady := TRUE;
			SetDiagOutput(i_etDiag := GD.ET_Diag.OK, i_etDiagExt := PDL_ET_DiagExt.WaitForStart, i_sMsg := '');
			diState := 5;
		END_IF
	END_IF
ELSIF NOT i_xEnable AND xEnableFlag THEN
	// detect negative flank on i_xEnable if FB is active
	fbHalt(Execute := FALSE);
	fbSetPos(Execute := FALSE);
	fbAbortTouchprobe(Execute := FALSE);
	fbTouchProbe(Execute := FALSE);
	fbMoveAbsolute(Execute := FALSE);
	fbMoveRelative(Execute := FALSE);
	xEnableFlag := FALSE;
	q_xReady    := FALSE;
	fbLoggerPoint.AddLogEntry(
		i_etLogLevel := APL.ET_LogLevel.UserAction, i_etDiag := q_etDiag, i_udiDiagExt := q_etDiagExt, i_sMessage := 'disable function block'
	);
	IF (diState <= 10) THEN
		// job not started yet -> disable immediately
		q_xActive    := FALSE;
		q_lrPosition := 0.0;
		q_xHomeOk    := FALSE;

		THIS^.SetDiagOutput(i_etDiag := GD.ET_Diag.Ok, i_etDiagExt := PDL_ET_DiagExt.Disabled, i_sMsg := '');
		diState := 0;
	ELSE
		// stop process before disable
		fbStop(Execute := TRUE);
		THIS^.SetDiagOutput(i_etDiag := GD.ET_Diag.Ok, i_etDiagExt := PDL_ET_DiagExt.WaitUntilDisabled, i_sMsg := '');
		diState := 100;
	END_IF
END_IF

IF q_xActive AND (i_ifDrive <> 0) THEN
	IF i_ifDrive.etAxisState < MOIN.ET_AxisState.Standstill AND diState > 0 AND diState < 100 THEN
		q_xMotionInstructionActive := FALSE;
		SetDiagOutput(
			i_etDiag    := GD.ET_Diag.DriveConditionInvalid,
			i_etDiagExt := PDL_ET_DiagExt.DriveNotReady,
			i_sMsg 		:= STANDARD.CONCAT(sDriveName,': AxisState < Standstill')
		);
		diState := 0;
	ELSIF i_ifDrive.etAxisState > MOIN.ET_AxisState.Stopping THEN
		xMotionJobStarted := TRUE; // latch a started job in order to make shure job has stared if for job finish is checked. This can be necessary if FB is called twice in a cycle as it is done in tests.
	END_IF
	q_lrPosition := i_ifDrive.RefPosition;
	(* The HW limits are evaluated depending on the mode – they must be queried during motion. *)
	IF i_etMode = PDL_ET_HomeTpMode.PosDirectionPosEdgeTp OR i_etMode = PDL_ET_HomeTpMode.PosDirectionNegEdgeTp THEN (* pos. direction *)
		xLimitGivenDirection    := i_xHWLimitPos;
		xLimitOpposideDirection := i_xHWLimitNeg;
	ELSE (* neg. direction *)
		xLimitGivenDirection    := i_xHWLimitNeg;
		xLimitOpposideDirection := i_xHWLimitPos;
	END_IF
END_IF

// statemachine of FB
CASE diState OF
	0: // FB is disabled or in error
		; // do nothing (error quit is done by negative flank of i_xEnable)

	5: 		fbAbortTouchprobe(Execute := TRUE);
			IF fbAbortTouchprobe.Done THEN
				fbAbortTouchprobe(Execute := FALSE);
				diState := 10;
			ELSIF fbAbortTouchprobe.Error THEN
				SetDiagOutput(
					i_etDiag    := GD.ET_Diag.UnexpectedProgramBehavior,
					i_etDiagExt := PDL_ET_DiagExt.UnexpectedFeedback,
					i_sMsg      := CONCAT('MC_AbortTrigger: ', PLCO.FC_EtResultToString(fbAbortTouchprobe.ErrorId))
				);
				diState := 0;
			END_IF

	10: // wait for start
		IF i_xStart THEN
			fbLoggerPoint.AddLogEntry(
				i_etLogLevel := APL.ET_LogLevel.UserAction, i_etDiag := q_etDiag, i_udiDiagExt := q_etDiagExt, i_sMessage := 'start function block'
			);
			q_xHomeOk := FALSE;
			IF NOT THIS^.StartParameterCheck() THEN
				// error during start (error message is already set during StartParameterCheck() )
				diState := 0;
			ELSE
				// store information of limit switches if search started on opposide limit switch in order to prevent error message from check of limit switches till run free from switch
				xLimitGivenDirectionOld    := xLimitGivenDirection;
				xLimitOpposideDirectionOld := xLimitOpposideDirection;
				// check all possible start conditions
				IF
					xLimitGivenDirection OR
					(NOT i_xRotativeSystem AND
						ifTouprobeData.Value AND
						(i_etMode = PDL_ET_HomeTpMode.PosDirectionPosEdgeTp OR i_etMode = PDL_ET_HomeTpMode.NegDirectionPosEdgeTp)) OR
					(NOT i_xRotativeSystem AND
						NOT ifTouprobeData.Value AND
						(i_etMode = PDL_ET_HomeTpMode.PosDirectionNegEdgeTp OR i_etMode = PDL_ET_HomeTpMode.NegDirectionNegEdgeTp))
				THEN
					// Standing on TP or not possible to drive in set direction -> search TP in different direction
					SetTpEdge(i_xOppositeFlank := TRUE);
					StartPositioningAndTPEdge(i_xOppositeDirection := TRUE);
					IF q_etDiag <> GD.ET_Diag.Ok THEN
						// exception during command, diag message already set in SearchTpInDifferentDirection()
						q_xMotionInstructionActive := FALSE;
						diState                    := 0;
					ELSE
						SetDiagOutput(i_etDiag := GD.ET_Diag.OK, i_etDiagExt := PDL_ET_DiagExt.WaitForNegEdgeOfTouchProbe, i_sMsg := '');
						diState := 40;
					END_IF
				ELSE
					// regular search of TP
					xLimitOpposideDirectionOld := xLimitOpposideDirection;
					SetTpEdge(i_xOppositeFlank := FALSE);
					StartPositioningAndTPEdge(i_xOppositeDirection := FALSE);
					IF q_etDiag <> GD.ET_Diag.Ok THEN
						// exception during command, diag message already set in SearchTpInDifferentDirection()
						q_xMotionInstructionActive := FALSE;
						diState                    := 0;
					ELSE
						IF xLimitOpposideDirection THEN
							SetDiagOutput(i_etDiag := GD.ET_Diag.Ok, i_etDiagExt := PDL_ET_DiagExt.WaitUntilLimitSwitchFree, i_sMsg := '');
						ELSE
							SetDiagOutput(i_etDiag := GD.ET_Diag.Ok, i_etDiagExt := PDL_ET_DiagExt.WaitForTouchProbeSignal, i_sMsg := '');
						END_IF
						diState := 20;
					END_IF
				END_IF
			END_IF
		END_IF
	20: // search TP in given direction
		fbMoveRelative(Execute := TRUE);
		IF ifTouprobeData.CaptureOk THEN
			fbMoveRelative(Execute := FALSE);
			fbLoggerPoint.AddLogEntry(
				i_etLogLevel := APL.ET_LogLevel.ExternalEvent,
				i_etDiag     := q_etDiag,
				i_udiDiagExt := q_etDiagExt,
				i_sMessage   := 'Touch probe found in given direction'
			);
			xMotionJobStarted  := FALSE;
			i_ifDrive.xIsHomed := TRUE;
			fbMoveAbsolute(Execute := TRUE, Position := ifTouprobeData.CaptureValue + i_lrOffset);

			IF fbMoveAbsolute.Error THEN
				SetDiagOutput(
					i_etDiag    := GD.ET_Diag.UnexpectedProgramBehavior,
					i_etDiagExt := PDL_ET_DiagExt.UnexpectedFeedback,
					i_sMsg      := CONCAT('MC_MoveAbsolute.ErrorID: ', PLCO.FC_EtResultToString(THIS^.fbMoveAbsolute.ErrorID))
				);
				fbMoveAbsolute(Execute := FALSE);
				diState := 0;
			ELSE
				q_xMotionInstructionActive := TRUE;
				// additional information after TP until offset is reached
				SetDiagOutput(i_etDiag := GD.ET_Diag.Ok, i_etDiagExt := PDL_ET_DiagExt.WaitForSensorSignal, i_sMsg := 'Offset movement in progress');

				diState := 60;
			END_IF
		ELSIF xLimitOpposideDirection AND NOT xLimitOpposideDirectionOld THEN
			fbStop(Execute := TRUE);
			fbMoveRelative(Execute := FALSE);
			IF i_etMode = PDL_ET_HomeTpMode.PosDirectionPosEdgeTp OR i_etMode = PDL_ET_HomeTpMode.PosDirectionNegEdgeTp THEN (* pos. direction *)
				SetDiagOutput(i_etDiag := GD.ET_Diag.LimitReached, i_etDiagExt := PDL_ET_DiagExt.HwLimitNegReached, i_sMsg := '');
			ELSE (* neg. direction *)
				SetDiagOutput(i_etDiag := GD.ET_Diag.LimitReached, i_etDiagExt := PDL_ET_DiagExt.HwLimitPosReached, i_sMsg := '');
			END_IF
			diState := 100;
		ELSIF xLimitGivenDirection AND NOT xLimitGivenDirectionOld THEN (* positive HW LimitSwitch *)
			fbMoveRelative(Execute := FALSE);
			fbLoggerPoint.AddLogEntry(
				i_etLogLevel := APL.ET_LogLevel.ExternalEvent,
				i_etDiag     := q_etDiag,
				i_udiDiagExt := q_etDiagExt,
				i_sMessage   := 'Limit switch in given direction seen'
			);
			fbHalt(Execute := TRUE);
			fbAbortTouchprobe(Execute := TRUE, Axis := i_ifDrive);
			IF fbAbortTouchprobe.Error THEN
				q_xMotionInstructionActive := FALSE;
				SetDiagOutput(
					i_etDiag    := GD.ET_Diag.UnexpectedProgramBehavior,
					i_etDiagExt := PDL_ET_DiagExt.UnexpectedFeedback,
					i_sMsg      := CONCAT('MC_AbortTrigger: ', PLCO.FC_EtResultToString(fbAbortTouchprobe.ErrorId))
				);
				fbAbortTouchprobe(Execute := FALSE);
				diState := 0;
			ELSE
				SetDiagOutput(i_etDiag := GD.ET_Diag.Ok, i_etDiagExt := PDL_ET_DiagExt.WaitUntilStopped, i_sMsg := '');
				diState := 30;
			END_IF
		ELSIF THIS^.fbMoveRelative.Done AND xMotionJobStarted THEN // positioning job for search of TP finisched
			THIS^.fbMoveRelative(Execute := FALSE);
			q_xMotionInstructionActive := FALSE;
			IF q_etDiagExt = PDL_ET_DiagExt.WaitUntilLimitSwitchFree THEN
				// give special exception message if the search started on limit switch and the limit switch was never set to false
				IF (i_etMode = PDL_ET_HomeTpMode.PosDirectionNegEdgeTp OR i_etMode = PDL_ET_HomeTpMode.PosDirectionPosEdgeTp) THEN
					SetDiagOutput(i_etDiag := GD.ET_Diag.HomingFailed, i_etDiagExt := PDL_ET_DiagExt.HwLimitNegStillActive, i_sMsg := '');
				ELSE
					SetDiagOutput(i_etDiag := GD.ET_Diag.HomingFailed, i_etDiagExt := PDL_ET_DiagExt.HwLimitPosStillActive, i_sMsg := '');
				END_IF
			ELSE
				SetDiagOutput(i_etDiag := GD.ET_Diag.HomingFailed, i_etDiagExt := PDL_ET_DiagExt.TouchProbeNotFound, i_sMsg := '');
			END_IF
			diState := 0;
		ELSIF NOT xLimitOpposideDirection AND xLimitOpposideDirectionOld THEN
			// signal user that the limit switch is left, which was active at start
			SetDiagOutput(i_etDiag := GD.ET_Diag.Ok, i_etDiagExt := PDL_ET_DiagExt.WaitForTouchProbeSignal, i_sMsg := '');
		ELSIF fbMoveRelative.Error THEN
			SetDiagOutput(
				i_etDiag    := GD.ET_Diag.UnexpectedProgramBehavior,
				i_etDiagExt := PDL_ET_DiagExt.UnexpectedFeedback,
				i_sMsg      := CONCAT('MC_MoveRelative.ErrorID: ', PLCO.FC_EtResultToString(THIS^.fbMoveRelative.ErrorID))
			);
			THIS^.fbMoveRelative(Execute := FALSE);
			diState := 0;
		END_IF
		xLimitGivenDirectionOld    := xLimitGivenDirection;
		xLimitOpposideDirectionOld := xLimitOpposideDirection;
	30: // wait until stopped after HW Limit reached during search in given direction
		fbAbortTouchprobe(Execute := TRUE);
		IF i_ifDrive.etAxisState <= MOIN.ET_AxisState.Standstill AND fbAbortTouchprobe.Done THEN
			fbAbortTouchprobe(Execute := FALSE);
			q_xMotionInstructionActive := FALSE;
			xLimitGivenDirection       := xLimitGivenDirectionOld;
			xLimitOpposideDirection    := xLimitOpposideDirectionOld;
			fbHalt(Execute := FALSE);
			SetTpEdge(i_xOppositeFlank := TRUE);
			StartPositioningAndTPEdge(i_xOppositeDirection := TRUE);
			IF q_etDiag <> GD.ET_Diag.Ok THEN
				// exception during command, diag message already set in SearchTpInDifferentDirection()
				q_xMotionInstructionActive := FALSE;
				diState                    := 0;
			ELSE
				SetDiagOutput(i_etDiag := GD.ET_Diag.OK, i_etDiagExt := PDL_ET_DiagExt.WaitForNegEdgeOfTouchProbe, i_sMsg := '');
				diState := 40;
			END_IF
		ELSIF fbAbortTouchprobe.Error THEN
				SetDiagOutput(
					i_etDiag    := GD.ET_Diag.UnexpectedProgramBehavior,
					i_etDiagExt := PDL_ET_DiagExt.UnexpectedFeedback,
					i_sMsg      := CONCAT('MC_AbortTrigger: ', PLCO.FC_EtResultToString(fbAbortTouchprobe.ErrorId))
				);
				fbAbortTouchprobe(Execute := FALSE);
				diState := 0;
		END_IF
	40: // search TP in opposite direction
		fbMoveRelative(Execute := TRUE);
		IF ifTouprobeData.CaptureOK = TRUE THEN
			fbLoggerPoint.AddLogEntry(
				i_etLogLevel := APL.ET_LogLevel.ExternalEvent,
				i_etDiag     := q_etDiag,
				i_udiDiagExt := q_etDiagExt,
				i_sMessage   := 'Touch probe found in opposite direction'
			);
			fbMoveRelative(Execute := FALSE);
			fbHalt(Execute := TRUE);
			SetDiagOutput(i_etDiag := GD.ET_Diag.OK, i_etDiagExt := PDL_ET_DiagExt.WaitUntilStopped, i_sMsg := '');
			diState := 50;

		ELSIF xLimitOpposideDirection AND NOT xLimitOpposideDirectionOld THEN // limit in opposite direction reached -> no more ways to searche TP
			fbMoveRelative(Execute := FALSE);
			fbStop(Execute := TRUE);
			IF i_etMode = PDL_ET_HomeTpMode.PosDirectionPosEdgeTp OR i_etMode = PDL_ET_HomeTpMode.PosDirectionNegEdgeTp THEN
				SetDiagOutput(i_etDiag := GD.ET_Diag.LimitReached, i_etDiagExt := PDL_ET_DiagExt.HwLimitNegReached, i_sMsg := '');
			ELSE (* neg. direction *)
				SetDiagOutput(i_etDiag := GD.ET_Diag.LimitReached, i_etDiagExt := PDL_ET_DiagExt.HwLimitPosReached, i_sMsg := '');
			END_IF
			diState := 100;

		ELSIF fbMoveRelative.Done AND xMotionJobStarted THEN // positioning has finished without finding TP or LimitSwitch
			q_xMotionInstructionActive := FALSE;
			SetDiagOutput(i_etDiag := GD.ET_Diag.HomingFailed, i_etDiagExt := PDL_ET_DiagExt.TouchProbeNotFound, i_sMsg := '');
			diState := 0;
		ELSIF fbMoveRelative.Error THEN
			SetDiagOutput(
				i_etDiag    := GD.ET_Diag.UnexpectedProgramBehavior,
				i_etDiagExt := PDL_ET_DiagExt.UnexpectedFeedback,
				i_sMsg      := CONCAT('MC_MoveRelative.ErrorID: ', PLCO.FC_EtResultToString(THIS^.fbMoveRelative.ErrorID))
			);
			THIS^.fbMoveRelative(Execute := FALSE);
			diState := 0;
		END_IF
		xLimitOpposideDirectionOld := xLimitOpposideDirection; // reset flag if not on sensor in order to detect error if sensor gets true again
		xLimitGivenDirectionOld    := xLimitGivenDirection;
	50: // whait Until Drive has stopped after finding TP in opposite direction
		fbHalt(Execute := TRUE);
		IF fbHalt.Done THEN
			fbHalt(Execute := FALSE);
			IF xLimitGivenDirection THEN
				q_xMotionInstructionActive := FALSE;
				IF i_etMode = PDL_ET_HomeTpMode.PosDirectionPosEdgeTp OR i_etMode = PDL_ET_HomeTpMode.PosDirectionNegEdgeTp THEN (* pos. direction *)
					SetDiagOutput(i_etDiag := GD.ET_Diag.LimitReached, i_etDiagExt := PDL_ET_DiagExt.HwLimitPosReached, i_sMsg := '');
				ELSE (* neg. direction *)
					SetDiagOutput(i_etDiag := GD.ET_Diag.LimitReached, i_etDiagExt := PDL_ET_DiagExt.HwLimitNegReached, i_sMsg := '');
				END_IF
				diState := 0;
			ELSE
				xLimitGivenDirectionOld    := xLimitGivenDirection;
				xLimitOpposideDirectionOld := xLimitOpposideDirection;
				SetTpEdge(i_xOppositeFlank := FALSE);
				StartPositioningAndTPEdge(i_xOppositeDirection := FALSE);
				IF q_etDiag <> GD.ET_Diag.Ok THEN
					// exception during command, diag message already set in StartPositioningAndTPEdge()
					q_xMotionInstructionActive := FALSE;
					diState                    := 0;
				ELSE
					SetDiagOutput(i_etDiag := GD.ET_Diag.Ok, i_etDiagExt := PDL_ET_DiagExt.WaitForTouchProbeSignal, i_sMsg := '');
					diState := 20;
				END_IF
			END_IF
		ELSIF fbHalt.Error THEN
			SetDiagOutput(
				i_etDiag    := GD.ET_Diag.UnexpectedProgramBehavior,
				i_etDiagExt := PDL_ET_DiagExt.UnexpectedFeedback,
				i_sMsg      := CONCAT('MC_Halt.ErrorID: ', PLCO.FC_EtResultToString(THIS^.fbHalt.ErrorID))
			);
			THIS^.fbHalt(Execute := FALSE);
			diState := 0;
		END_IF
	60: // wait till positioning done after seen TP
		fbMoveAbsolute(Execute := TRUE);
		IF fbMoveAbsolute.Done THEN // pos finished
			fbMoveAbsolute(Execute := FALSE);
			q_xMotionInstructionActive := FALSE;
			fbSetPos(Execute := TRUE, Relative := FALSE, Position := i_lrHomePosition);
			IF fbSetPos.Error THEN
				SetDiagOutput(
					i_etDiag    := GD.ET_Diag.UnexpectedProgramBehavior,
					i_etDiagExt := PDL_ET_DiagExt.UnexpectedFeedback,
					i_sMsg      := CONCAT('MC_Setpos: ', PLCO.FC_EtResultToString(fbSetPos.ErrorId))
				);
				fbSetPos(Execute := FALSE);
				diState := 0;
			ELSE
				fbSetPos(Execute := FALSE);
				q_xHomeOk := TRUE;
				SetDiagOutput(i_etDiag := GD.ET_Diag.Ok, i_etDiagExt := PDL_ET_DiagExt.HomingDone, i_sMsg := '');
				IF NOT i_xStart THEN
					diState := 10;
				ELSE
					diState := 70;
				END_IF
			END_IF
		ELSIF fbMoveAbsolute.Error THEN
			SetDiagOutput(
				i_etDiag    := GD.ET_Diag.UnexpectedProgramBehavior,
				i_etDiagExt := PDL_ET_DiagExt.UnexpectedFeedback,
				i_sMsg      := CONCAT('MC_MoveAbsolute.ErrorID: ', PLCO.FC_EtResultToString(THIS^.fbMoveAbsolute.ErrorID))
			);
			THIS^.fbMoveAbsolute(Execute := FALSE);
			q_xMotionInstructionActive := FALSE;
			diState                    := 0;
		END_IF
	70: // wait till i_xStart FALSE to prevent immediate restart
		IF NOT i_xStart THEN
			fbLoggerPoint.AddLogEntry(
				i_etLogLevel := APL.ET_LogLevel.DebugMessage, i_etDiag := q_etDiag, i_udiDiagExt := q_etDiagExt, i_sMessage := 'i_xStart reset'
			);
			// diagnosis output keeps ET_Diag.Ok and PDL_ET_DiagExt.HomingDone as it is set in state 60
			diState := 10;
		END_IF
	100: // wait  until stopped after HW Limit and Error
		fbStop(Execute := TRUE);
		IF
			i_ifDrive.etAxisState = MOIN.ET_AxisState.Disabled OR
			i_ifDrive.etAxisState = MOIN.ET_AxisState.ErrorStop OR
			i_ifDrive.etAxisState = MOIN.ET_AxisState.Standstill OR
			fbStop.Done
		THEN
			q_xMotionInstructionActive := FALSE;
			fbStop(Execute := FALSE);
			fbLoggerPoint.AddLogEntry(
				i_etLogLevel := APL.ET_LogLevel.DebugMessage, i_etDiag := q_etDiag, i_udiDiagExt := q_etDiagExt, i_sMessage := 'Axis stopped'
			);

			IF NOT xEnableFlag THEN
				q_xActive    := FALSE;
				q_lrPosition := 0.0;
				q_xHomeOk    := FALSE;
				SetDiagOutput(i_etDiag := GD.ET_Diag.OK, i_etDiagExt := PDL_ET_DiagExt.Disabled, i_sMsg := '');
			END_IF

			diState := 0;
		END_IF

		IF fbStop.Error AND fbStop.ErrorId <> PLCO.ET_Result.StoppingInterrupted THEN
			q_xMotionInstructionActive := FALSE;
			q_xReady                   := FALSE;
			SetDiagOutput(
				i_etDiag    := GD.ET_Diag.UnexpectedProgramBehavior,
				i_etDiagExt := PDL_ET_DiagExt.UnexpectedFeedback,
				i_sMsg      := CONCAT('MC_Stop.ErrorID:', PLCO.FC_EtResultToString(fbStop.ErrorId))
			);
			fbStop(Execute := FALSE);
			diState := 0;
		END_IF
	ELSE
		q_xReady := FALSE;
		THIS^.SetDiagOutput(
			i_etDiag := GD.ET_Diag.UnexpectedProgramBehavior, i_etDiagExt := PDL_ET_DiagExt.UnknownState, i_sMsg := DINT_TO_STRING(diState)
		);
		diState := 0;
END_CASE

(* ---- PDL_FB_MovingAverage.fb.st ---- *)
{attribute 'no_explicit_call' := 'Do not call body of FB_Average'}
FUNCTION_BLOCK PDL_FB_MovingAverage

VAR
	uiOrder_loc			: UINT := 1;

	lrAverage_loc		: LREAL;
	xInitialized		: BOOL;

	uiI					: UINT;
	uiLevel_loc			: UINT;
	uiWriteIndex		: UINT;
	alrBufferElements	: ARRAY[1..Gc_uiMovingAverageMaxOrder] OF LREAL;

	lrSum				: LREAL;
	uiValidValues		: UINT;
END_VAR

;

(* ---- PDL_FB_PosIn.fb.st ---- *)
FUNCTION_BLOCK PDL_FB_PosIn
VAR_INPUT
	i_ifDrive        : Moin.IF_Axis;
	i_xSensor        : BOOL;
	i_xPosEdge       : BOOL;
	i_lrMaxTravel    : LREAL;
	i_lrOffset       : LREAL;
	i_lrVelocity     : LREAL;
	i_lrAcceleration : LREAL;
	i_lrDeceleration : LREAL;
	i_lrJerk         : LREAL;
	i_xStart         : BOOL;
END_VAR
VAR_OUTPUT
	q_xError          : BOOL;
	q_diErrorId       : PLCO.ET_Result;
	q_xInOk           : BOOL;
	q_xSensorNotFound : BOOL;
	q_xMoveToHomePosition: BOOL;

END_VAR
VAR
	diState        : DINT;
	xPosEdgeFlag   : BOOL;
	xNegEdgeFlag   : BOOL;
	xTPFlag        : BOOL;
	fbMoveRelative : PLCO.MC_MoveRelative;
	fbMoveRelativeOffset : PLCO.MC_MoveRelative;
END_VAR

IF i_xStart = TRUE THEN
	q_xINOk           := FALSE;
	q_xSensorNotFound := FALSE;
	q_xError          := FALSE;
	q_diErrorId       := PLCO.ET_Result.Ok;
	q_xMoveToHomePosition := FALSE;
	xPosEdgeFlag      := FALSE;
	xNegEdgeFlag      := FALSE;
	xTPFlag           := i_xSensor;
	diState           := 10;
	THIS^.fbMoveRelative(Execute := FALSE);
	THIS^.fbMoveRelativeOffset(Execute := FALSE);
END_IF

IF i_xSensor AND NOT xTPFlag THEN
	xTPFlag      := TRUE;
	xPosEdgeFlag := TRUE;
ELSIF NOT i_xSensor AND xTPFlag THEN
	xTPFlag      := FALSE;
	xNegEdgeFlag := TRUE;
END_IF

CASE diState OF

	0: (*Fertig *)
		THIS^.fbMoveRelative(Execute := FALSE);
		THIS^.fbMoveRelativeOffset(Execute := FALSE);

	10: (* PosStart *)
		THIS^.fbMoveRelative(
			Axis         := i_ifDrive,
			Execute      := TRUE,
			Distance     := i_lrMaxTravel,
			Velocity     := i_lrVelocity,
			Acceleration := i_lrAcceleration,
			Deceleration := i_lrDeceleration,
			Jerk         := i_lrJerk,
			BufferMode   := PLCO.MC_Buffer_Mode.Aborting);

		IF THIS^.fbMoveRelative.Error THEN
			q_xError    := TRUE;
			q_diErrorId := THIS^.fbMoveRelative.ErrorId;
			diState := 0;
		ELSE
			diState := 30;
		END_IF

	30: (* Warten bis TP gesehen *)
		THIS^.fbMoveRelative();

		IF THIS^.fbMoveRelative.Error THEN
			q_xError    := TRUE;
			q_diErrorId := THIS^.fbMoveRelative.ErrorId;
			diState := 0;

		ELSIF (i_xPosEdge AND xPosEdgeFlag) OR (NOT i_xPosEdge AND xNegEdgeFlag) THEN
			THIS^.fbMoveRelative(Execute := FALSE);

			THIS^.fbMoveRelativeOffset(
				Axis         := i_ifDrive,
				Execute      := TRUE,
				Distance     := i_lrOffset,
				Velocity     := i_lrVelocity,
				Acceleration := i_lrAcceleration,
				Deceleration := i_lrDeceleration,
				Jerk         := i_lrJerk,
				BufferMode   := PLCO.MC_Buffer_Mode.Aborting);

			IF THIS^.fbMoveRelativeOffset.Error THEN
				q_xError    := TRUE;
				q_diErrorId := THIS^.fbMoveRelativeOffset.ErrorId;
				diState := 0;
			ELSE
				q_xMoveToHomePosition := TRUE;
				diState := 50;
			END_IF

		ELSIF THIS^.fbMoveRelative.Error THEN
			q_xError    := TRUE;
			q_diErrorId := THIS^.fbMoveRelative.ErrorId;
			diState := 0;

		ELSIF THIS^.fbMoveRelative.Done THEN (* maxTravel zu Ende *)
			q_xSensorNotFound := TRUE;
			diState           := 0;
		END_IF

	50: (* Warten bis steht *)
		THIS^.fbMoveRelativeOffset();
		IF THIS^.fbMoveRelativeOffset.Done THEN
			q_xINOk    := TRUE;
			diState    := 0;

		ELSIF THIS^.fbMoveRelativeOffset.Error THEN
			q_xError    := TRUE;
			q_diErrorId := THIS^.fbMoveRelativeOffset.ErrorId;
			diState := 0;
		END_IF

END_CASE

(* ---- PDL_FB_ResetTrackingDeviation.fb.st ---- *)
FUNCTION_BLOCK PDL_FB_ResetTrackingDeviation IMPLEMENTS SE_Async.IF_Async
VAR_INPUT
END_VAR
VAR_OUTPUT
END_VAR
VAR
	xDone_loc                   : BOOL;
	ifDrive2_loc                : DDI.IF_Drive2;
	lrOldTrackingDeviationLimit : LREAL;
END_VAR

(* ---- PDL_FB_SetDrvEncPos.fb.st ---- *)
FUNCTION_BLOCK PDL_FB_SetDrvEncPos IMPLEMENTS SE_Async.IF_Async
VAR_INPUT
END_VAR
VAR_OUTPUT
END_VAR
VAR
	ifDeviceType_loc 		: DeviceTypeInterfaces.IF_Device_Type;
	diResultSetDrvEnc_loc	: DINT;
	lrPosition_loc			: LREAL;
	xDone_loc				: BOOL;
END_VAR

(* ---- PDL_FB_SetDrvEncPosGetState.fb.st ---- *)
FUNCTION_BLOCK PDL_FB_SetDrvEncPosGetState IMPLEMENTS SE_Async.IF_Async
VAR_INPUT
END_VAR
VAR_OUTPUT
END_VAR
VAR
	ifDeviceType_loc 		: DeviceTypeInterfaces.IF_Device_Type;
	diResultSetDrvEncGetState_loc	: DINT;
	xDone_loc						: BOOL;
END_VAR

(* ---- PDL_FB_SetTrackingDeviation.fb.st ---- *)
FUNCTION_BLOCK PDL_FB_SetTrackingDeviation IMPLEMENTS SE_Async.IF_Async
VAR_INPUT
END_VAR
VAR_OUTPUT
END_VAR
VAR
	xDone_loc                       : BOOL;
	ifDrive2_loc                    : DDI.IF_Drive2;
	lrOldTrackingDeviationLimit     : LREAL;
	lrCurrentTrackingDeviationLimit : LREAL;
END_VAR

(* ---- PDL_FB_WriteDriveEncoder.fb.st ---- *)
FUNCTION_BLOCK PDL_FB_WriteDriveEncoder
VAR_INPUT
	i_xEnable        : BOOL;
	i_ifDrive        : MOIN.IF_Axis;
	i_lrHomePos      : LREAL;
	i_lrAbsEncOffset : LREAL;
	i_lrUserPeriod   : LREAL;
	i_xExecute       : BOOL;
END_VAR

VAR_OUTPUT
	q_xActive   : BOOL;
	q_xReady    : BOOL;
	q_xBusy     : BOOL;
	q_xDone     : BOOL;
	q_etDiag    : GD.ET_Diag     := GD.ET_Diag.OK;
	q_etDiagExt : PDL_ET_DiagExt := PDL_ET_DiagExt.Disabled;
	q_sMsg      : STRING[80];
END_VAR

VAR CONSTANT
	c_lrStandStillVel : LREAL := 10.0;
	c_timDisableTime  : TIME  := T#1500MS;
	c_timProgramTime  : TIME  := T#1000MS;
	c_lrRealNull      : LREAL := 10E-12;
END_VAR
VAR
	ifScalingAccess        : DMFI.IF_ScalingAccess;
	ifScaling              : DMFI.IF_Scaling;
	ifDrive2Access         : DDI.IF_Drive2Access;
	ifDrive2               : DDI.IF_Drive2;
	ifDriveConfigAccess    : DDI.IF_DriveConfigAccess;
	ifDriveConfig          : DDI.IF_DriveConfig;
	ifDriveAccess          : DMFI.IF_DriveAccess;
	ifDrive                : DMFI.IF_Drive;
	ifMotorAccess          : DDI.IF_MotorAccess;
	ifMotor                : DDI.IF_Motor;
	ifEncoderAccess        : DDI.IF_EncoderAccess;
	ifEncoder              : DDI.IF_Encoder;
	ifLXM62DriveAccess     : LXM62SI.IF_Lexium62DriveAccess;
	ifLXM62Drive           : LXM62SI.IF_Lexium62Drive;
	ifWorkingModeAccess    : CFDI.IF_WorkingModeAccess;
	ifWorkingMode          : CFDI.IF_WorkingMode;
	ifDeviceType		   : DeviceTypeInterfaces.IF_Device_Type;
	xSuccess               : BOOL;
	xInterfacesInitialised : BOOL;

	xEnableFlag : BOOL;

	diResult         : DINT;
	diState          : DINT;
	lrEncoderPeriode : LREAL;
	lrSavePosition   : LREAL;
	tonTimeOut       : Standard.TON;
	diSercosState    : DINT;
	uiI              : UINT;
	lrSum            : LREAL;
	lrAverage        : LREAL;
	alrA             : ARRAY[0..17] OF LREAL;
	xValid           : BOOL;
	lrModuloPosition : LREAL;
	xAxisEnableFlag  : BOOL;

	lrEncoderRange : LREAL;
	etDiag         : GD.ET_Diag;
	etDiagExt      : PDL_ET_DiagExt;

	fbSetDrvEncPos         : PDL_FB_SetDrvEncPos;
	fbSetDrvEncPosGetState : PDL_FB_SetDrvEncPosGetState;
	lrPositionTemp         : LREAL;
	diWritePositionState   : DINT;
	xError                 : BOOL;
	etResult               : SE_Async.ET_Result;
	sResultMsg             : STRING(80);
	fbPower                : PLCO.MC_Power;
	sMsg                   : STRING(80);
END_VAR

IF i_xEnable AND NOT xEnableFlag THEN (* Pos. edge on i_xExecute *)
	xEnableFlag := TRUE;

	q_xActive := TRUE;
	q_xReady  := FALSE;
	q_xDone   := FALSE;

	SetDiagOutput(i_etDiag := GD.ET_Diag.OK, i_etDiagExt := PDL_ET_DiagExt.Initializing, i_sMsg := '');

	diState := 0;

	xInterfacesInitialised := FALSE;

	IF ParameterCheckEnable() THEN
		xInterfacesInitialised := TRUE;

		IF SE_Async.G_ifAsyncMgr.xInitDone THEN
			q_xReady := TRUE;
			SetDiagOutput(i_etDiag := GD.ET_Diag.OK, i_etDiagExt := PDL_ET_DiagExt.WaitForExecute, i_sMsg := '');
			diState := 5;
		ELSE
			SE_Async.G_ifAsyncMgr.Init();
			diState := 150;
		END_IF
	END_IF

ELSIF NOT i_xEnable AND xEnableFlag THEN (* Neg. edge on Enable *)
	xEnableFlag := FALSE;

	xInterfacesInitialised := FALSE;

	q_xActive := FALSE;
	q_xReady  := FALSE;
	q_xBusy   := FALSE;
	q_xDone   := FALSE;

	SetDiagOutput(i_etDiag := GD.ET_Diag.OK, i_etDiagExt := PDL_ET_DiagExt.Disabled, i_sMsg := '');
	diState := 0;

ELSIF NOT q_xActive THEN
	RETURN;
END_IF

IF xInterfacesInitialised THEN
	AverageVel();
	q_xBusy := q_etDiag = GD.ET_Diag.Ok AND NOT q_xDone AND diState > 5;
END_IF

CASE diState OF

	-1000:
		IF fbSetDrvEncPosGetState.xDone THEN
			diState := 21;
		END_IF
	-1003:
		SE_Async.G_ifAsyncMgr.Init(q_xError => xError, q_etResult => etResult, q_sResultMsg => sResultMsg);
		IF xError THEN
			AsyncExtDiagTranslation(i_etResult := etResult);
			diState := 0;
		ELSIF SE_Async.G_ifAsyncMgr.xInitDone THEN
			q_xReady := TRUE;
			SetDiagOutput(i_etDiag := GD.ET_Diag.Ok, i_etDiagExt := PDL_ET_DiagExt.WaitForExecute, i_sMsg := '');
			diState := 5;
		END_IF
	0: (* Idle or Error *)
		;
	5:
		IF i_xExecute THEN

			lrSavePosition  := i_ifDrive.RefPosition; (* Save Axis Position *)
			xAxisEnableFlag := i_ifDrive.etAxisState >= MOIN.ET_AxisState.Standstill; (* Save state of Axis *)
			//fb needs a edge therefore calling fb twice
			fbPower(Axis := i_ifDrive, Enable := TRUE);
			fbPower(Axis := i_ifDrive, Enable := FALSE);

			tonTimeOut(IN := FALSE, PT := c_timDisableTime);
			xValid := FALSE;

			FOR uiI := 1 TO 16 DO (* delete array of AverageVel() *)
				alrA[uiI] := 0;
			END_FOR

			uiI   := 1;
			lrSum := 0;

			SetDiagOutput(i_etDiag := GD.ET_Diag.OK, i_etDiagExt := PDL_ET_DiagExt.WaitUntilDriveDisabled, i_sMsg := '');
			diState := 6;
		END_IF
	6:
		tonTimeOut(IN := TRUE);

		IF tonTimeOut.Q THEN
			diState := 10;
		END_IF
	10: (* Waiting for axis disabled *)

		(* Timeout for disabling axis and axis not standing *)
		IF (ABS(lrAverage) >= c_lrStandStillVel) THEN
			q_xReady := FALSE;

			SetDiagOutput(i_etDiag := GD.ET_Diag.DriveConditionInvalid, i_etDiagExt := PDL_ET_DiagExt.DriveIsMoving, i_sMsg := '');
			diState := 0;

			(* Timeout for disabling axis and axis not disabled*)
		ELSIF i_ifDrive.etAxisState > MOIN.ET_AxisState.Disabled THEN
			q_xReady := FALSE;

			SetDiagOutput(i_etDiag := GD.ET_Diag.DriveConditionInvalid, i_etDiagExt := PDL_ET_DiagExt.DriveNotDisabled, i_sMsg := '');

			diState := 0;

			(* Timeout for disabling axis and axis is disabled and standing*)
		ELSIF (ABS(lrAverage) < c_lrStandStillVel) THEN
			diState              := 11; // 	WritePosition();
			diWritePositionState := 10;
		END_IF
	11:
		WritePosition();
	20: (* Wait for programming done *)
		tonTimeOut(IN := TRUE);
		(* Writing time over *)
		IF tonTimeOut.Q THEN
			fbSetDrvEncPosGetState.ifDeviceType := ifDeviceType;
			SE_Async.G_ifAsyncMgr.Start(i_ifAsync := fbSetDrvEncPosGetState, q_etResult => etResult, q_sResultMsg => sResultMsg, q_xError => xError);

			IF xError THEN
				AsyncExtDiagTranslation(i_etResult := etResult);
				RETURN;
			ELSE
				diState := -1000;
			END_IF
		END_IF
	21:
		diResult := fbSetDrvEncPosGetState.diResultSetDrvEncGetState;
		IF diResult = 0 THEN

			PDL_FC_ReadDriveEncoder(
				i_ifDrive        := i_ifDrive, (* Read Position from Encoder *)
				i_lrHomePos      := i_lrHomePos,
				i_lrAbsEncOffset := i_lrAbsEncOffset,
				i_lrUserPeriod   := i_lrUserPeriod,
				q_etDiag         => etDiag,
				q_etDiagExt      => etDiagExt,
				q_sMsg			 => sMsg
			);

			IF etDiag <> GD.ET_Diag.Ok THEN
				q_xReady := FALSE;

				SetDiagOutput(
					i_etDiag    := GD.ET_Diag.UnexpectedProgramBehavior,
					i_etDiagExt := PDL_ET_DiagExt.UnexpectedFeedback,
					i_sMsg      := CONCAT('FC_ReadDriveEncoder: ', UDINT_TO_STRING(etDiagExt))
				);

				diState := 0;
				RETURN;
			END_IF

			IF xAxisEnableFlag THEN (* Restore original State *)
				//fb needs a edge therefore calling fb twice
				fbPower(Axis := i_ifDrive, Enable := FALSE);
				fbPower(Axis := i_ifDrive, Enable := TRUE);
				IF fbPower.Error THEN
					q_xReady := FALSE;

					SetDiagOutput(
						i_etDiag    := GD.ET_Diag.UnexpectedProgramBehavior,
						i_etDiagExt := PDL_ET_DiagExt.UnexpectedFeedback,
						i_sMsg      := CONCAT('fbPower: ', TO_STRING(fbPower.ErrorId))
					);

					diState := 0;
					RETURN;
				END_IF

				SetDiagOutput(i_etDiag := GD.ET_Diag.Ok, i_etDiagExt := PDL_ET_DiagExt.WaitUntilDriveEnabled, i_sMsg := '');
				diState := 30;
			ELSE
				q_xDone := TRUE;

				SetDiagOutput(i_etDiag := GD.ET_Diag.Ok, i_etDiagExt := PDL_ET_DiagExt.WritingPositionDone, i_sMsg := '');

				diState := 0;
			END_IF

		ELSIF diResult = 2 THEN
			q_xReady := FALSE;

			SetDiagOutput(i_etDiag := GD.ET_Diag.DriveConditionInvalid, i_etDiagExt := PDL_ET_DiagExt.ProgrammingInvalidEEPROM, i_sMsg := '');
			diState := 0;

		ELSIF diResult = 3 THEN
			q_xReady := FALSE;

			SetDiagOutput(i_etDiag := GD.ET_Diag.DriveConditionInvalid, i_etDiagExt := PDL_ET_DiagExt.NoAccessToEEPROM, i_sMsg := '');
			diState := 0;

		ELSE
			q_xReady := FALSE;

			SetDiagOutput(i_etDiag := GD.ET_Diag.UnexpectedProgramBehavior, i_etDiagExt := PDL_ET_DiagExt.EncoderWriteTimeOut, i_sMsg := '');
			diState := 0;
		END_IF
	30: (* Wait for AxisState => standstill *)
		IF i_ifDrive.etAxisState >= MOIN.ET_AxisState.Standstill THEN
			q_xDone := TRUE;

			SetDiagOutput(i_etDiag := GD.ET_Diag.Ok, i_etDiagExt := PDL_ET_DiagExt.WritingPositionDone, i_sMsg := '');

			diState := 0;
		END_IF

		(* End of case *)
	ELSE
		q_xReady := FALSE;

		SetDiagOutput(
			i_etDiag := GD.ET_Diag.UnexpectedProgramBehavior, i_etDiagExt := PDL_ET_DiagExt.UnknownState, i_sMsg := DINT_TO_STRING(diState)
		);
		diState := 0;
END_CASE
